(* IEC 61131-3 sources: llm-plc-st-eval/data/definitivo/gemini-3.1-pro-preview/C8/few_shot, 3 files *)

(* ---- ejec_1.st ---- *)
FUNCTION_BLOCK FB_Valvula
VAR_INPUT
    nivelAlto : BOOL; (* Contacto NA que inicia el temporizador *)
END_VAR
VAR_OUTPUT
    valvula : BOOL; (* Bobina de salida *)
END_VAR
VAR
    T1 : TON; (* Temporizador a la conexión *)
END_VAR

(* Rama 1: El contacto nivelAlto alimenta la entrada IN del temporizador T1 *)
T1(IN := nivelAlto, PT := T#5S);

(* Rama 2: El contacto NA de T1.Q alimenta la bobina valvula *)
valvula := T1.Q;
END_FUNCTION_BLOCK

(* ---- ejec_2.st ---- *)
FUNCTION_BLOCK FB_Valvula
VAR_INPUT
    nivelAlto : BOOL; (* Contacto NA que inicia el temporizador *)
END_VAR
VAR_OUTPUT
    valvula : BOOL; (* Bobina activada por el temporizador *)
END_VAR
VAR
    T1 : TON; (* Temporizador a la conexion *)
END_VAR

(* Rama 1: Llamada al temporizador TON con PT de 5 segundos *)
T1(IN := nivelAlto, PT := T#5S);

(* Rama 2: La bobina se activa con la salida Q del temporizador *)
valvula := T1.Q;
END_FUNCTION_BLOCK

(* ---- ejec_3.st ---- *)
FUNCTION_BLOCK FB_Valvula
VAR_INPUT
    nivelAlto : BOOL; (* Contacto NA que activa el temporizador *)
END_VAR
VAR_OUTPUT
    valvula : BOOL; (* Bobina de salida *)
END_VAR
VAR
    T1 : TON; (* Temporizador a la conexion *)
END_VAR

(* Rama 1: El contacto alimenta la entrada IN del temporizador TON *)
T1(IN := nivelAlto, PT := T#5S);

(* Rama 2: El contacto de la salida del temporizador alimenta la bobina *)
valvula := T1.Q;
END_FUNCTION_BLOCK
